(* IEC 61131-3 sources: T4Exjobb/Sigma/Stations/Terminal/HMI/Network/LseRtkAlarm, 1 file *)

(* ---- ONE_LseRtkAlarm_Table.st ---- *)
#define OBJECTS_CONFIG

#include "..\..\Class\_AlarmX0Para\_AlarmX0Para.h"
#include <.\lsl_st_mt.h>
#include "..\..\Class\_AlarmXBuffer\AlarmXBuffer.h"

FUNCTION GLOBAL TAB ONE_LseRtkAlarm
-1$UINT, 0$UINT,
0$UINT, 0$UINT,

3$UDINT,
TO_UDINT(800276940), "_AlarmX0Para", 0$UINT, 11$UINT, 1$UINT,
TO_UDINT(315844732), "_AlarmX1Para", 0$UINT, 2$UINT, 1$UINT,
TO_UDINT(2835625764), "_AlarmXBuffer", 0$UINT, 19$UINT, 1$UINT,

_NO_ATTR, TO_UDINT(3323358457), "EMERGENCYSTOP",

_NO_ATTR, TO_UDINT(108736354), "SERVERERROR",

_NO_ATTR, TO_UDINT(3212185425), "_ALARMXBUFFER1",

//Internal connections
0$UDINT,
0$UDINT,
0$UDINT,
0$UDINT,

//Initialization values
0$UDINT,
3$UDINT,
TO_UDINT(0), "Config", TO_UDINT(1),//|LseRtkAlarm.EmergencyStop.Config;
TO_UDINT(1), "Config", TO_UDINT(2),//|LseRtkAlarm.ServerError.Config;
TO_UDINT(2), "No", TO_UDINT(64),//|LseRtkAlarm._AlarmXBuffer1.No;

//Symbolic initialization values
0$UDINT,
0$UDINT,

//Initialization of string values
0$UDINT,
0$UDINT,

//Configuration of tasks (RealTime, Cyclic, Background)
0$UDINT,
0$UDINT,

0$UDINT,
0$UDINT,

0$UDINT,
0$UDINT,

//External connections
0$UDINT,
0$UDINT,

//Magic internal connections
0$UDINT,
0$UDINT,

//Configuration of timeslots of tasks (RealTime, Cyclic)
#ifdef __LSLLDR_TIMESLOTS__
0$UDINT,
0$UDINT,

0$UDINT,
0$UDINT,

#endif //__LSLLDR_TIMESLOTS__

//MultiMaster connections
#ifdef __LSLLDR_MULTIMASTER__
0$UDINT,
0$UDINT,
#endif //__LSLLDR_MULTIMASTER__

//Configuration for task ID (RealTime, CyclicTime)
#ifdef __LSLLDR_TASKID__
"\\\\TASKS2  "
0$UDINT,
0$UDINT,

0$UDINT,
0$UDINT,

0$UDINT,
0$UDINT,

#endif //__LSLLDR_TASKID__

END_FUNCTION
